(* IEC 61131-3 sources: llm-plc-st-eval/data/definitivo/claude-sonnet-4-6/B1/zero_shot, 3 files *)

(* ---- ejec_1.st ---- *)
```pascal
FUNCTION_BLOCK FB_Motor
VAR_INPUT
    btnMarcha : BOOL; (* Botón de marcha: TRUE = pulsado *)
    btnParo   : BOOL; (* Botón de paro: TRUE = pulsado *)
    btnEmerg  : BOOL; (* Paro de emergencia: TRUE = activado *)
END_VAR

VAR_OUTPUT
    motorOn : BOOL; (* Salida al contactor del motor *)
END_VAR

VAR
    bloqueado : BOOL; (* Enclavamiento por emergencia *)
END_VAR

(*
    Lógica de control:
    - btnParo y btnEmerg se asumen como contacto normalmente cerrado
      representado en lógica positiva: TRUE = fallo/paro activo.
    - bloqueado se activa con btnEmerg y solo se resetea manualmente
      (aquí se mantiene hasta un ciclo sin emergencia Y sin marcha,
       o bien puede requerir un reset explícito según la aplicación).
    - Para rearrancar tras emergencia se debe soltar btnEmerg
      y NO tener btnMarcha activo en ese mismo ciclo (reset seguro).
*)

(* 1. Activar enclavamiento si se detecta emergencia *)
IF btnEmerg THEN
    bloqueado := TRUE;
END_IF;

(* 2. Reset del enclavamiento: solo cuando NO hay emergencia
      Y NO hay botón de marcha pulsado (evita rearranque automático) *)
IF NOT btnEmerg AND NOT btnMarcha THEN
    bloqueado := FALSE;
END_IF;

(* 3. Lógica de marcha/paro con auto-retención (seal-in) *)
IF btnEmerg OR btnParo OR bloqueado THEN
    (* Paro prioritario: emergencia, paro normal o enclavamiento activo *)
    motorOn := FALSE;
ELSIF btnMarcha THEN
    (* Arranque: flanco o nivel, el motor se enciende *)
    motorOn := TRUE;
END_IF;
(* Si ninguna condición aplica, motorOn conserva su valor anterior
   → auto-retención implementada por la variable de salida misma *)

END_FUNCTION_BLOCK
```

(* ---- ejec_2.st ---- *)
```pascal
FUNCTION_BLOCK FB_Motor
VAR_INPUT
    btnMarcha : BOOL; (* Botón de marcha: TRUE = pulsado *)
    btnParo   : BOOL; (* Botón de paro: TRUE = pulsado *)
    btnEmerg  : BOOL; (* Paro de emergencia: TRUE = activado *)
END_VAR

VAR_OUTPUT
    motorOn : BOOL; (* Salida al contactor del motor *)
END_VAR

VAR
    bloqueado : BOOL; (* Enclavamiento por emergencia *)
END_VAR

(*
    Lógica de control:
    1. Si se activa la emergencia → parar motor y bloquear rearranque.
    2. Si se pulsa paro → parar motor (sin bloqueo).
    3. Si se pulsa marcha Y no hay bloqueo → arrancar motor (set).
    4. El motor se mantiene encendido por auto-retención (motorOn se conserva).
*)

(* --- Gestión del enclavamiento por emergencia --- *)
IF btnEmerg THEN
    bloqueado := TRUE;  (* Bloqueo permanente hasta reset manual *)
END_IF;

(* --- Paro: emergencia o botón de paro --- *)
IF btnEmerg OR btnParo THEN
    motorOn := FALSE;

(* --- Arranque: marcha pulsada, sin bloqueo y sin paro activo --- *)
ELSIF btnMarcha AND NOT bloqueado THEN
    motorOn := TRUE;

(* --- Auto-retención: si no hay orden nueva, mantener estado actual --- *)
(* (motorOn conserva su valor al no asignarse en otra rama) *)
END_IF;
```

(* ---- ejec_3.st ---- *)
```pascal
FUNCTION_BLOCK FB_Motor
VAR_INPUT
    btnMarcha : BOOL; (* Botón de marcha: TRUE = pulsado *)
    btnParo   : BOOL; (* Botón de paro: TRUE = pulsado *)
    btnEmerg  : BOOL; (* Paro de emergencia: TRUE = activado *)
END_VAR

VAR_OUTPUT
    motorOn : BOOL; (* Salida al contactor del motor *)
END_VAR

VAR
    bloqueado : BOOL; (* Enclavamiento por emergencia *)
END_VAR

(*
    Lógica de control:
    1. Si se activa la emergencia → parar motor y bloquear rearranque.
    2. Si se pulsa paro → parar motor (sin bloqueo).
    3. Si está bloqueado → no permitir arranque aunque btnMarcha esté activo.
    4. Si se pulsa marcha y no hay bloqueo ni paro → arrancar y retener (automantenimiento).
*)

(* --- Gestión del enclavamiento por emergencia --- *)
IF btnEmerg THEN
    bloqueado := TRUE;  (* Activa bloqueo; solo un reset manual lo limpia *)
END_IF;

(* --- Lógica de paro con prioridad sobre marcha --- *)
IF btnEmerg OR btnParo THEN
    motorOn := FALSE;   (* Paro inmediato en cualquier caso *)

(* --- Lógica de arranque: solo si no hay bloqueo activo --- *)
ELSIF btnMarcha AND NOT bloqueado THEN
    motorOn := TRUE;    (* Arranque + automantenimiento por la propia salida *)
END_IF;

(* Nota: el automantenimiento lo garantiza el PLC al conservar el valor
   de motorOn entre ciclos; no se necesita contacto auxiliar explícito
   en ST porque la variable retiene su estado hasta que se modifique. *)
```

---

### Explicación de la lógica

| Condición | `bloqueado` | `motorOn` |
|---|---|---|
| `btnEmerg` = TRUE | Se pone TRUE | FALSE |
| `btnParo` = TRUE | Sin cambio | FALSE |
| `btnMarcha` = TRUE y `bloqueado` = FALSE | Sin cambio | TRUE |
| `btnMarcha` = TRUE y `bloqueado` = TRUE | Sin cambio | Permanece FALSE |
| Ningún botón pulsado | Sin cambio | Retiene estado anterior |

> **Reset del enclavamiento:** la variable `bloqueado` se mantiene en `TRUE` hasta que un procedimiento externo (p. ej. un reset supervisado) la ponga a `FALSE`. Esto cumple el requisito de que tras un paro de emergencia el motor **no rearranque** aunque `btnMarcha` siga activo.
